FUNCTION_BLOCK INIT2 (* E_TRIG Counterpart, Stufe 2 (E2Init) *)
  (* Standard: 61131-3; Classification: standard boolean function; Description: Copyright (c) 2011 TU Wien ACIN, HR Agrartechnik GmbH This program and the accompanying materials are made available under the terms of the Eclipse Public License 2.0 which is available at https://www.eclipse.org/legal/epl-2.0/ SPDX-License-Identifier: EPL-2.0 *)
  (* Version 3.2, 2026-10-30, Franz Höpfinger, Meisterschulen am Ostbahnhof, INIT-Stufe 2: nach dem App-INIT (EInit). E_TRIG mit EVENTTYPE E2Init loest den unverbundenen Eingang aus, INIT2O an das INIT des Ziels. *)
  (* Version 3.1, 2026-10-11, Franz Höpfinger, Meisterschulen am Ostbahnhof, Organization-Attribut ergaenzt (XSD-Pflichtfeld). Basis fuer die neue INIT_ON/INIT_OFF/INIT_ON_OFF-Familie (eigenstaendige EInitOn/EInitOff Pass-Through-Kanaele). *)
  (* Version 3.0, 2025-04-14, Patrick Aigner, Eclipse 4diac, changed package *)
  (* Version 1.0, 2011-06-21, Monika Wenger, TU Wien ACIN, initial API and implementation and/or initial documentation *)
  PACKAGE events::init;
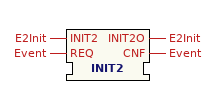
  EVENT_INPUT
    INIT2 : E2Init; (* Initialization Request *)
    REQ; (* Service Request *)
  END_EVENT
  EVENT_OUTPUT
    INIT2O : E2Init; (* Initialization Confirm *)
    CNF; (* Confirmation of Requested Service *)
  END_EVENT
  EVENT_CONNECTIONS
    INIT2 TO INIT2O;
    REQ TO CNF;
  END_CONNECTIONS
END_FUNCTION_BLOCK
